// TIA Portal V19 export
DATA_BLOCK "ALL_VALVES_DB"   // DB3
// stored: InstanceOfName ALL_VALVES, InstanceOfType FB
"ALL_VALVES"
   // VAR
   //    XV01 { S7_SetPoint := 'True'} : "valve";
   //    XV02 { S7_SetPoint := 'True'} : "valve";
   //    XV03 { S7_SetPoint := 'True'} : "valve";
   //    XV04 { S7_SetPoint := 'True'} : "valve";
   //    XV05 { S7_SetPoint := 'True'} : "valve";
   //    XV06 { S7_SetPoint := 'True'} : "valve";
   //    XV07 { S7_SetPoint := 'True'} : "valve";
   //    XV08 { S7_SetPoint := 'True'} : "valve";
   // END_VAR
BEGIN
END_DATA_BLOCK
